SUBAPPLICATION NumericValue_TO_AUI2 (* VT-Eingabefeld (CInputNumber) lesen und als AUI2 (bidirektional) an einen Consumer weiterreichen (z.B. AOption_AUI_DEMUX_N.K). Speichert NICHT selbst - der Consumer meldet den tatsaechlich uebernommenen Wert ueber denselben AUI2-Plug zurueck, das Echo wird auf das VT-Feld zurueckgeschrieben. *)
  (* Standard: 61499-2; Description: Copyright (c) 2026 Meisterschulen am Ostbahnhof This program and the accompanying materials are made available under the terms of the Eclipse Public License 2.0 which is available at https://www.eclipse.org/legal/epl-2.0/ SPDX-License-Identifier: EPL-2.0 *)
  (* Version 1.0, 2026-10-13, Franz Höpfinger, Meisterschulen am Ostbahnhof, Ausgelagert aus Uebung_094c_AX (dort je Dropdown inline dupliziert: NumericValue_IDA+AD_TO_AUI+AUI_TO_AUI2+AUI_TO_AUDI+Q_NumericValue_AUDI) zur Wiederverwendung. Analog MyLib::sys::NumericValue_TO_AR2, aber UINT/AUI2 statt REAL/AR2 und einfaches u16ObjId statt stObj (kein Scale/Offset/Decimals fuer einen reinen Index-Wert noetig). *)
  PACKAGE MyLib::sys;
  IMPORT isobus::UT::Q::const::IDs::ID_NULL;
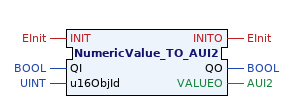
  EVENT_INPUT
    INIT : EInit; (* Initialization Request *)
  END_EVENT
  EVENT_OUTPUT
    INITO : EInit; (* Initialization Confirm *)
  END_EVENT
  VAR_INPUT
    QI : BOOL := TRUE; (* Quality Input - TRUE to enable service *)
    u16ObjId : UINT := ID_NULL; (* Object ID *)
  END_VAR
  VAR_OUTPUT
    QO : BOOL; (* Quality Output - TRUE if service executed successfully *)
  END_VAR
  PLUGS
    VALUEO : adapter::types::bidirectional::AUI2;
  END_PLUGS
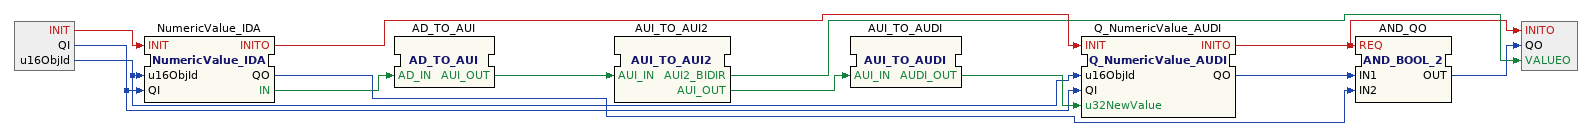
  FBS
    NumericValue_IDA : isobus::UT::io::NumericValue::NumericValue_IDA;
    AD_TO_AUI : adapter::conversion::unidirectional::AD_TO_AUI;
    AUI_TO_AUI2 : adapter::conversion::bidirectional::AUI_TO_AUI2;
    AUI_TO_AUDI : adapter::conversion::unidirectional::AUI_TO_AUDI;
    Q_NumericValue_AUDI : isobus::UT::Q::Q_NumericValue_AUDI;
    AND_QO : iec61131::booleanOperators::AND_BOOL_2;
  END_FBS
  EVENT_CONNECTIONS
    INIT TO NumericValue_IDA.INIT;
    NumericValue_IDA.INITO TO Q_NumericValue_AUDI.INIT;
    Q_NumericValue_AUDI.INITO TO INITO;
    Q_NumericValue_AUDI.INITO TO AND_QO.REQ;
  END_CONNECTIONS
  DATA_CONNECTIONS
    u16ObjId TO NumericValue_IDA.u16ObjId;
    u16ObjId TO Q_NumericValue_AUDI.u16ObjId;
    QI TO Q_NumericValue_AUDI.QI;
    QI TO NumericValue_IDA.QI;
    Q_NumericValue_AUDI.QO TO AND_QO.IN1;
    NumericValue_IDA.QO TO AND_QO.IN2;
    AND_QO.OUT TO QO;
  END_CONNECTIONS
  ADAPTER_CONNECTIONS
    NumericValue_IDA.IN TO AD_TO_AUI.AD_IN;
    AD_TO_AUI.AUI_OUT TO AUI_TO_AUI2.AUI_IN;
    AUI_TO_AUI2.AUI2_BIDIR TO VALUEO;
    AUI_TO_AUI2.AUI_OUT TO AUI_TO_AUDI.AUI_IN;
    AUI_TO_AUDI.AUDI_OUT TO Q_NumericValue_AUDI.u32NewValue;
  END_CONNECTIONS
END_SUBAPPLICATION
